FUNCTION_BLOCK TcoKukaKss_StopMovementsTask_v_9_3_x EXTENDS TcoKukaKssTask_v_9_3_x
VAR
	_stopType : TcoAbstractions.eTcoRoboticsStopType;
END_VAR

IF Execute() THEN
	_blink(inOnTime:=T#500MS,inOffTime:=T#500MS);

	IF _progress = 0 THEN
		IF CheckReferences() THEN
			_progress := _progress + 1;
		END_IF
	END_IF

	IF _progress = 1 THEN
		// AX step 0: waiting for 'RobotStopped'
		inoControl.MoveEnable := FALSE;
		_varInfo :=__VARINFO(inoStatus.State.RobotStopped);
		THIS^.Messenger.OnCondition(_infoTimer.Q AND NOT inoStatus.State.RobotStopped).Warning(_sb.Clear().Append('<#Waiting for signal: #>').Append(_varInfo.Symbol).ToString());
		IF inoStatus.State.RobotStopped THEN
			_progress := _progress + 1;
		END_IF
	END_IF

	IF _progress = 2 THEN
		DoneWhen(TRUE);
	END_IF

	CallTimers(TRUE);
	THIS^.ThrowWhen(_errorTimer.Q);
END_IF

IF THIS^.Error AND NOT _errorMessage.Pinned THEN
	THIS^.Restore();
END_IF

METHOD INTERNAL InvokeWithParams : ITcoTaskStatus
VAR_INPUT
	inStopType : eTcoRoboticsStopType;
END_VAR
_stopType := inStopType;
InvokeWithParams := THIS^.Invoke();
END_METHOD

METHOD PUBLIC FB_init : BOOL
VAR_INPUT
    bInitRetains : BOOL; // if TRUE, the retain variables are initialized (warm start / cold start)
    bInCopyCode : BOOL; // if TRUE, the instance afterwards gets moved into the copy code (online change)
    ParentObject : ITcoObject;
END_VAR
END_METHOD

(*~
	<docu>
		<summary>
			Executes when task is aborted.
		</summary>			
	</docu>	
~*)
METHOD PROTECTED OnAbort
IF __ISVALIDREF(inoStatus) THEN THIS^.inoStatus.ActionDescription := '<#Stop movements was aborted.#>'; END_IF;
END_METHOD

(*~
	<docu>
		<summary>
			Executes when task reaches the ```Done``` state .
		</summary>			
	</docu>	
~*)
METHOD PROTECTED OnDone
IF __ISVALIDREF(inoStatus) THEN THIS^.inoStatus.ActionDescription := '<#Stop movements finished successfully.#>'; END_IF;
_progress := 0;
END_METHOD

(*~
	<docu>
		<summary>
			Executes when task reaches the ```Error``` state.
		</summary>			
	</docu>	
~*)
METHOD PROTECTED OnError
VAR
	description: STRING;
END_VAR
description := '<#Stop movements finished with error.#>';
IF __ISVALIDREF(inoStatus) THEN THIS^.inoStatus.ActionDescription := description; END_IF;
THIS^._errorMessage.Error(_sb.Clear().Append(description).Append(' To restore acknowledge this alarm.').ToString()).Pin();
END_METHOD

METHOD PROTECTED OnStart
IF __ISVALIDREF(inoStatus) THEN THIS^.inoStatus.ActionDescription := '<#Stop movements started.#>'; END_IF;
CallTimers(FALSE);
END_METHOD

(*~
	<docu>
		<summary>
			Restores this instance to the Ready state. Can be called explicitly or from within one of the restore mechanisms.
			<para>
				See also <see cref="PlcDocu.TcoCore.TcoTask.AutoRestorable()"/>
			</para>
		</summary>
	</docu>
~*)
METHOD Restore : ITcoRestorable
SUPER^.Restore();
END_METHOD

END_FUNCTION_BLOCK

(* stored: Version 1.1.0.1, ProductVersion 3.1.4024.12
   POU TcoKukaKss_StopMovementsTask_v_9_3_x: Id {f92d8be1-c95b-45f3-b6ea-93b7aa49e2c0}, SpecialFunc None
   Method InvokeWithParams: Id {90e1d21f-2fdd-45e2-b8bb-47356c40529d}
   Method FB_init: Id {109fb7ae-b18c-4ca8-a155-adc8318097a5}
   Method OnAbort: Id {c3265f02-64e2-474d-893c-b0fea90f61fa}
   Method OnDone: Id {1426ea81-35fc-48a9-a9c7-7f842a491e53}
   Method OnError: Id {c897726c-ea27-4e53-9528-edded7c9c9c7}
   Method OnStart: Id {fe655c4a-103f-4552-a164-3c5620bc81d7}
   Method Restore: Id {c229f1ab-6dc4-4be9-ae18-008f2aad404d} *)
